Fanuc KAREL source: KO00123.KL

PROGRAM KO00123
%NOLOCKGROUP
VAR
  A: ARRAY[2] OF SHORT
  B: REAL
  OUT: INTEGER
BEGIN
  A[1] = 1
  B = 2
  OUT = ATAN2(A[1], B)
END KO00123
